    rq_activate_all_grippers(True)
    # end: URCap Program Node
  end
  $ 59 "zero_ftsensor()"
  zero_ftsensor()
  $ 60 "EXTT"
  $ 61 "Set GRP_3F_Enable=Off"
  set_standard_digital_out(4, False)
  $ 62 "Set DO[6]=Off"
  set_standard_digital_out(6, False)
  $ 63 "Set GRP_3F_Decap=Off"
  set_standard_digital_out(3, False)
  $ 64 "Set GRP_3F_Cap=Off"
  set_standard_digital_out(2, False)
  $ 65 "Set GRP_3F_Open=Off"
  set_standard_digital_out(5, False)
  $ 66 "PSE_T≔get_tool_free_pose(dir=[0,0,0.150], move_in_base_frame=True)"
  global PSE_T=get_tool_free_pose(dir=[0,0,0.150], move_in_base_frame=True)
  $ 67 "If is_reachable(Base_const, [PSE_T])"
  if (is_reachable(p[0.0,0.0,0.0,0.0,0.0,0.0], [PSE_T])):
    $ 68 "MoveL"
    $ 69 "PSE_T" "breakAfter"
    movel(PSE_T, a=1.2, v=0.15)
  end
  $ 70 "powder dispensing variable init"
  $ 71 "Start_thread≔ False "
  global Start_thread=  False
  $ 72 "vib_mot_thread≔ False "
  global vib_mot_thread=  False
  $ 73 "kp≔0.00005"
  global kp=0.00005
  $ 74 "ki≔0.0005"
  global ki=0.0005
  $ 75 "kd≔0.002"
  global kd=0.002
  $ 76 "dt≔0.02"
  global dt=0.02
  $ 77 "Integral_error≔0"
  global Integral_error=0
  $ 78 "current_error≔0"
  global current_error=0
  $ 79 "previous_error≔0"
  global previous_error=0
  $ 80 "tilt_increment≔0"
  global tilt_increment=0
  $ 81 "tilt_angle≔0"
  global tilt_angle=0
  $ 82 "diff≔0"
  global diff=0
  $ 83 "current_pose≔get_actual_tcp_pose()"
  global current_pose= get_actual_tcp_pose ()
  $ 84 "Relative_trans≔p[0, 0, -0.035, 0, 0, 0]"
  global Relative_trans=p[0, 0, -0.035, 0, 0, 0]
  $ 85 "ContA_plc_offst≔p[-0.00205, 0.02547, 0.03730, -0.03, -2.183, 6.165]"
  global ContA_plc_offst=p[-0.00205, 0.02547, 0.03730, -0.03, -2.183, 6.165]
  $ 86 "PowA_50_offset≔p[0.21808, -0.19943, 0.06584, 0, 0, 0]"
  global PowA_50_offset=p[0.21808, -0.19943, 0.06584, 0, 0, 0]
  $ 87 "scooping_init()"
  scooping_init()
  $ 88 "tilt_init_reference()"
  tilt_init_reference()
  $ 89 "switch_spatula≔ True "
  global switch_spatula=  True
  $ 679 "Thread_1"
  thread Thread_1():
    while (True):
      $ 680 "If Start_thread≟ True "
      if (Start_thread ==   True  ):
        $ 681 "Weight_value≔get_weight()"
        global Weight_value=get_weight()
        $ 682 "Wait: 0.1"
        sleep(0.1)
        $ 683 "sync()"
        sync()
      end
    end
  end
  threadId_Thread_1 = run Thread_1()
  $ 695 "Thread_2"
  thread Thread_2():
    while (True):
      $ 696 "Loop vib_mot_thread≟ True "
      thread Thread_while_696():
        while (True):
          $ 697 "diff≔Target_weight-Weight_value"
          global diff=Target_weight-Weight_value
          $ 698 "If diff>0.15"
          global thread_flag_698=0
          thread Thread_if_698():
            $ 700 "Set AO[0]=4.0"
            set_standard_analog_out(0, 0.4)
            thread_flag_698 = 1
          end
          if (diff>0.15):
            global thread_handler_698=run Thread_if_698()
            while (thread_flag_698 == 0):
              if not(diff>0.15):
                kill thread_handler_698
                thread_flag_698 = 2
              else:
                sync()
              end
            end
          else:
            thread_flag_698 = 2
          end
          if (thread_flag_698 == 2):
            $ 701 "ElseIf diff≥0.05 and diff≤0.15"
            global thread_flag_701=0
            thread Thread_if_701():
              $ 702 "vibration_2()"
              vibration_2()
              thread_flag_701 = 1
            end
            if (diff >= 0.05 and diff <= 0.15):
              global thread_handler_701=run Thread_if_701()
              while (thread_flag_701 == 0):
                if not(diff >= 0.05 and diff <= 0.15):
                  kill thread_handler_701
                  thread_flag_701 = 2
                else:
                  sync()
                end
              end
            else:
              thread_flag_701 = 2
            end
            if (thread_flag_701 == 2):
              $ 703 "ElseIf diff≥0.01 and diff<0.05"
              if (diff >= 0.01 and diff<0.05):
                $ 704 "vibration_3()"
                vibration_3()
              else:
                $ 705 "ElseIf diff>0 and diff<0.01"
                if (diff>0 and diff<0.01):
                  $ 706 "vibration_4()"
                  vibration_4()
                else:
                  $ 707 "Else" "noBreak"
                  $ 708 "Set AO[0]=0.0"
                  set_standard_analog_out(0, 0.0)
                end
              end
            end
          end
        end
      end
      if (vib_mot_thread ==   True  ):
        global thread_handler_696=run Thread_while_696()
        while (vib_mot_thread ==   True  ):
          sync()
        end
        kill thread_handler_696
      end
      $ 712 "sync()"
      sync()
    end
  end
  threadId_Thread_2 = run Thread_2()
  while (True):
    $ 90 "Robot Program"
    $ 91 "MAIN"
    $ 92 "command_manager(external_control='uGO', cond_suspend=(ITM_Manipulated and AMR_AtTarget and AMR_Charging and AMR_Battery<40), cond_unsuspend=(AMR_Battery≟60))"
    command_manager(external_control="uGO", cond_suspend=(ITM_Manipulated  and  AMR_AtTarget  and  AMR_Charging  and  AMR_Battery<40), cond_unsuspend=(AMR_Battery == 60))
    $ 93 "log_state(STATE_Info)"
    log_state(STATE_Info)
    $ 94 "Switch STATE"
    switch_1 = STATE
    $ 95 "Case 1"
    if (1 == switch_1):
      $ 96 "Stopping"
      $ 97 "STATE_Info≔'Stopping'"
      global STATE_Info="Stopping"
      $ 98 "end_freedrive_mode()"
      end_freedrive_mode()
      $ 99 "Set"
      set_tcp(p[0.0,0.0,0.161,3.1415,0.0,0.0])
      $ 100 "PSE_T≔get_tool_free_pose(dir=[0,0,0.150], move_in_base_frame=True)"
      global PSE_T=get_tool_free_pose(dir=[0,0,0.150], move_in_base_frame=True)
      $ 101 "If is_reachable(Base_const, [PSE_T])"
      if (is_reachable(p[0.0,0.0,0.0,0.0,0.0,0.0], [PSE_T])):
        $ 102 "MoveL"
        $ 103 "PSE_T" "breakAfter"
        movel(PSE_T, a=1.2, v=0.15)
      end
      $ 104 "do_transition(keep_rxry=OBJ_Picked, r=0)"
      do_transition(keep_rxry=OBJ_Picked, r=0)
      $ 113 "Call Sub_AMR_MiR_V3"
      Sub_AMR_MiR_V3()
      $ 114 "If stopping() and AMR_Done"
      if (stopping()  and  AMR_Done):
        $ 115 "STATE≔2"
        global STATE=2
        $ 116 "ugo_update_outputs()"
        ugo_update_outputs()
      end
    elif (2 == switch_1):
      $ 117 "Case 2"
      $ 118 "Stopped"
      $ 119 "STATE_Info≔'Stopped'"
      global STATE_Info="Stopped"
      $ 120 "Call Sub_AMR_MiR_V3"
      Sub_AMR_MiR_V3()
      $ 121 "If CMD_Reset"
      if (CMD_Reset):
        $ 122 "STATE≔3"
        global STATE=3
        $ 123 "ugo_update_outputs()"
        ugo_update_outputs()
      end
    elif (3 == switch_1):
      $ 124 "Case 3"
      $ 125 " Resetting"
      $ 126 "STATE_Info≔'Resetting'"
      global STATE_Info="Resetting"
      $ 127 "uML"
      $ 128 "reset_error()"
      reset_error()
      $ 129 "reset_warning()"
      reset_warning()
      $ 130 "PROCESS_Step≔0"
      global PROCESS_Step=0
      $ 131 "PROCESS_Info≔''"
      global PROCESS_Info=""
      $ 132 "ARM_Referenced≔ False "
      global ARM_Referenced=  False
      $ 133 "WRK_Done≔ False "
      global WRK_Done=  False
      $ 134 "ITM_Prepared≔ False "
      global ITM_Prepared=  False
      $ 135 "ITM_Manipulated≔ False "
      global ITM_Manipulated=  False
      $ 136 "STP≔0"
      global STP=0
      $ 137 "Action≔0"
      global Action=0
      $ 138 "Action_Info≔''"
      global Action_Info=""
      $ 139 "ITM_ID≔0"
      global ITM_ID=0
      $ 140 "JIG≔0"
      global JIG=0
      $ 141 "JIG_Slot≔0"
      global JIG_Slot=0
      $ 142 "Task_info≔''"
      global Task_info=""
      $ 143 "Set"
      set_tcp(p[0.0,0.0,0.161,3.1415,0.0,0.0])
      $ 144 "App"
      $ 145 "'ADD APPLICATION SPECIFIC COMMANDS'"
      # 'ADD APPLICATION SPECIFIC COMMANDS'
      $ 146 "OBJ_Type≔0"
      global OBJ_Type=0
      $ 147 "OBJ_Nbr≔0"
      global OBJ_Nbr=0
      $ 148 "If CNT_Rack_Output≥50"
      if (CNT_Rack_Output >= 50):
        $ 149 "CNT_Rack_Output≔0"
        global CNT_Rack_Output=0
      end
      $ 150 "TASK≔struct(ID=0, NAVI=struct(target=0, footprint=0, protectiveOff=0, dock=0), WORK=struct(ITM_ID_Src=0, JIG_ID_Src=0, OBJ_Nbr_Src=0, ACT_Src=0, ITM_ID_Tgt=0, JIG_ID_Tgt=0, OBJ_Nbr_Tgt=0, ACT_Tgt=0, OBJ_Type=0))"
      global TASK=struct(ID=0, NAVI=struct(target=0, footprint=0, protectiveOff=0, dock=0), WORK=struct(ITM_ID_Src=0, JIG_ID_Src=0, OBJ_Nbr_Src=0, ACT_Src=0, ITM_ID_Tgt=0, JIG_ID_Tgt=0, OBJ_Nbr_Tgt=0, ACT_Tgt=0, OBJ_Type=0))
      $ 151 "Call Sub_AMR_MiR_V3"
      Sub_AMR_MiR_V3()
      $ 152 "If resetting() and AMR_Done"
      if (resetting()  and  AMR_Done):
        $ 153 "STATE≔4"
        global STATE=4
        $ 154 "ugo_update_outputs()"
        ugo_update_outputs()
      end
    elif (4 == switch_1):
      $ 155 "Case 4"
      $ 156 "Idle"
      $ 157 "STATE_Info≔'Idle'"
      global STATE_Info="Idle"
      $ 158 "If CMD_Start"
      if (CMD_Start):
        $ 159 "STATE≔5"
        global STATE=5
        $ 160 "ugo_update_outputs()"
        ugo_update_outputs()
      end
    elif (5 == switch_1):
      $ 161 "Case 5"
      $ 162 "Starting"
      $ 163 "STATE_Info≔'Starting'"
      global STATE_Info="Starting"
      $ 164 "'ADD COMMANDS WHAT TO START WITH'"
      # 'ADD COMMANDS WHAT TO START WITH'
      $ 165 "Call Sub_AMR_MiR_V3"
      Sub_AMR_MiR_V3()
      $ 166 "get ugo data"
      $ 167 "Assign Tasks"
      $ 168 "TASK.ID = ugo_get_task()"
      TASK.ID = ugo_get_task()
      $ 169 "If TASK.ID≟1"
      if (TASK.ID == 1):
        $ 170 "Task_info≔'Charge'"
        global Task_info="Charge"
        $ 171 "Parameters"
        $ 172 "AMR_PosTarget≔1"
        global AMR_PosTarget=1
      else:
        $ 173 "ElseIf TASK.ID≟9"
        if (TASK.ID == 9):
          $ 174 "'Pick Sarstedt Rack from Variable source'"
          # 'Pick Sarstedt Rack from Variable source'
          $ 175 "Task_info≔'Navigate to Target'"
          global Task_info="Navigate to Target"
          $ 176 "Parameters"
          $ 177 "AMR_PosTarget≔UGO.read_input('00','ITM_ID')"
          global AMR_PosTarget=UGO.read_input("00","ITM_ID")
        else:
          $ 178 "ElseIf TASK.ID≟49"
          if (TASK.ID == 49):
            $ 179 "Task_info≔'Pick Containers'"
            global Task_info="Pick Containers"
            $ 180 "Parameters"
            $ 181 "ITM_ID≔1"
            global ITM_ID=1
            $ 182 "OBJ_Type≔6"
            global OBJ_Type=6
            $ 183 "JIG≔15"
            global JIG=15
            $ 184 "AMR_PosTarget≔3"
            global AMR_PosTarget=3
          else:
            $ 185 "ElseIf TASK.ID≟50"
            if (TASK.ID == 50):
              $ 186 "Task_info≔'Decap Containers'"
              global Task_info="Decap Containers"
              $ 187 "Parameters"
              $ 188 "ITM_ID≔1"
              global ITM_ID=1
              $ 189 "OBJ_Type≔6"
              global OBJ_Type=6
              $ 190 "JIG≔16"
              global JIG=16
              $ 191 "AMR_PosTarget≔5"
              global AMR_PosTarget=5
            else:
              $ 192 "ElseIf TASK.ID≟51"
              if (TASK.ID == 51):
                $ 193 "Task_info≔'Detect Spatula and transfer powder'"
                global Task_info="Detect Spatula and transfer powder"
                $ 194 "Parameters"
                $ 195 "ITM_ID≔1"
                global ITM_ID=1
                $ 196 "Target_weight≔(UGO.read_input('00','Target_weight'))/1000"
                global Target_weight=(UGO.read_input("00","Target_weight"))/1000
                $ 197 "OBJ_Type≔8"
                global OBJ_Type=8
                $ 198 "JIG≔16"
                global JIG=16
                $ 199 "AMR_PosTarget≔5"
                global AMR_PosTarget=5
              else:
                $ 200 "ElseIf TASK.ID≟52"
                if (TASK.ID == 52):
                  $ 201 "Task_info≔'Pick PowderA'"
                  global Task_info="Pick PowderA"
                  $ 202 "Parameters"
                  $ 203 "ITM_ID≔1"
                  global ITM_ID=1
                  $ 204 "OBJ_Type≔6"
                  global OBJ_Type=6
                  $ 205 "JIG≔15"
                  global JIG=15
                  $ 206 "AMR_PosTarget≔3"
                  global AMR_PosTarget=3
                else:
                  $ 207 "ElseIf TASK.ID≟53"
                  if (TASK.ID == 53):
                    $ 208 "Task_info≔'Decap PowderA'"
                    global Task_info="Decap PowderA"
                    $ 209 "Parameters"
                    $ 210 "ITM_ID≔1"
                    global ITM_ID=1
                    $ 211 "OBJ_Type≔6"
                    global OBJ_Type=6
                    $ 212 "JIG≔1"
                    global JIG=1
                    $ 213 "AMR_PosTarget≔5"
                    global AMR_PosTarget=5
                  else:
                    $ 214 "ElseIf TASK.ID≟54"
                    if (TASK.ID == 54):
                      $ 215 "Task_info≔'Dispense PowderA'"
                      global Task_info="Dispense PowderA"
                      $ 216 "Parameters"
                      $ 217 "ITM_ID≔1"
                      global ITM_ID=1
                      $ 218 "Target_weight≔(UGO.read_input('00','Target_weight'))/1000"
                      global Target_weight=(UGO.read_input("00","Target_weight"))/1000
                      $ 219 "W_now≔(UGO.read_input('00','Container_weight'))/1000"
                      global W_now=(UGO.read_input("00","Container_weight"))/1000
                      $ 220 "Powder_name≔(UGO.read_input('00','Powder_name'))"
                      global Powder_name=(UGO.read_input("00","Powder_name"))
                      $ 221 "OBJ_Type≔6"
                      global OBJ_Type=6
                      $ 222 "JIG≔17"
                      global JIG=17
                      $ 223 "AMR_PosTarget≔5"
                      global AMR_PosTarget=5
                    else:
                      $ 224 "ElseIf TASK.ID≟55"
                      if (TASK.ID == 55):
                        $ 225 "Task_info≔'Place PowderA'"
                        global Task_info="Place PowderA"
                        $ 226 "Parameters"
                        $ 227 "ITM_ID≔1"
                        global ITM_ID=1
                        $ 228 "OBJ_Type≔6"
                        global OBJ_Type=6
                        $ 229 "JIG≔21"
                        global JIG=21
                        $ 230 "AMR_PosTarget≔5"
                        global AMR_PosTarget=5
                      else:
                        $ 231 "Else" "noBreak"
                        $ 232 "set_error(ERROR_WRONG_ORDER)"
                        set_error(ERROR_WRONG_ORDER)
                      end
                    end
                  end
                end
              end
            end
          end
        end
      end
      $ 233 "test ugo"
      $ 234 "Wait: 0.2"
      sleep(0.2)
      $ 235 "ugo_update_outputs()"
      ugo_update_outputs()
      $ 236 "If starting() and AMR_Done"
      if (starting()  and  AMR_Done):
        $ 237 "log_message(Task_info, 'New Task: ')"
        log_message(Task_info, "New Task: ")
        $ 238 "log_message(to_str(TASK.ID), 'Task_ID: ')"
        log_message(to_str(TASK.ID), "Task_ID: ")
        $ 239 "do_transition(keep_rxry=OBJ_Picked)"
        do_transition(keep_rxry=OBJ_Picked)
        $ 240 "STATE≔6"
        global STATE=6
        $ 241 "ugo_update_outputs()"
        ugo_update_outputs()
      end
    elif (6 == switch_1):
      $ 242 "Case 6"
      $ 243 "Execute"
      $ 244 "STATE_Info≔'Execute'"
      global STATE_Info="Execute"
      $ 245 "If  not CMD_Hold and not CMD_Suspend"
      global thread_flag_245=0
      thread Thread_if_245():
        $ 246 "Switch PROCESS_Step"
        switch_2 = PROCESS_Step
        $ 247 "Case 0"
        if (0 == switch_2):
          $ 248 "PROCESS_Info≔'process control'"
          global PROCESS_Info="process control"
          $ 249 "log_process(PROCESS_Info)"
          log_process(PROCESS_Info)
          $ 250 "process control"
          $ 251 "If  not AMR_AtTarget"
          if (  not  AMR_AtTarget):
            $ 252 "PROCESS_Step≔1"
            global PROCESS_Step=1
          else:
            $ 253 "ElseIf (( not ITM_Prepared and  not WRK_Done) or (ITM_Prepared and WRK_Done))"
            if (((  not  ITM_Prepared  and    not  WRK_Done)  or  (ITM_Prepared  and  WRK_Done))):
              $ 254 "PROCESS_Step≔2"
              global PROCESS_Step=2
            else:
              $ 255 "ElseIf  not WRK_Done"
              if (  not  WRK_Done):
                $ 256 "PROCESS_Step≔3"
                global PROCESS_Step=3
              else:
                $ 257 "Else" "noBreak"
                $ 258 "task finished"
                $ 259 "PROCESS_Info≔''"
                global PROCESS_Info=""
                $ 260 "STATE≔7"
                global STATE=7
                $ 261 "ugo_update_outputs()"
                ugo_update_outputs()
              end
            end
          end
        elif (1 == switch_2):
          $ 262 "Case 1"
          $ 263 "navigate"
          $ 264 "'MOVING THE uML'"
          # 'MOVING THE uML'
          $ 265 "PROCESS_Info≔'move to target'"
          global PROCESS_Info="move to target"
          $ 266 "log_process(PROCESS_Info)"
          log_process(PROCESS_Info)
          $ 267 "If TASK.ID≟1"
          if (TASK.ID == 1):
            $ 268 "Action≔51"
            global Action=51
          else:
            $ 269 "Else" "noBreak"
            $ 270 "Action≔52"
            global Action=52
          end
          $ 271 "Call Sub_AMR_MiR_V3"
          Sub_AMR_MiR_V3()
          $ 272 "If AMR_Done"
          if (AMR_Done):
            $ 273 "PROCESS_Step≔0"
            global PROCESS_Step=0
          end
        elif (2 == switch_2):
          $ 274 "Case 2"
          $ 275 "prepare"
          $ 276 "'THINGS THAT HAVE TO BE DONE ONCE IN A SEQUENCE,WORKFLOW'"
          # 'THINGS THAT HAVE TO BE DONE ONCE IN A SEQUENCE,WORKFLOW'
          $ 277 "PROCESS_Info≔'prepare for work'"
          global PROCESS_Info="prepare for work"
          $ 278 "log_process(PROCESS_Info)"
          log_process(PROCESS_Info)
          $ 279 "If TASK.WORK.ITM_ID_Src>1"
          if (TASK.WORK.ITM_ID_Src>1):
            $ 280 "ITM_ID≔TASK.WORK.ITM_ID_Src"
            global ITM_ID=TASK.WORK.ITM_ID_Src
          else:
            $ 281 "ElseIf TASK.WORK.ITM_ID_Tgt>1"
            if (TASK.WORK.ITM_ID_Tgt>1):
              $ 282 "ITM_ID≔TASK.WORK.ITM_ID_Tgt"
              global ITM_ID=TASK.WORK.ITM_ID_Tgt
            end
          end
          $ 283 "If  not ARM_Referenced and (ITM_ID≠0)"
          if (  not  ARM_Referenced  and  (ITM_ID != 0)):
            $ 284 "STP≔1"
            global STP=1
          else:
            $ 285 "ElseIf ARM_Referenced or (ITM_ID≟0)"
            if (ARM_Referenced  or  (ITM_ID == 0)):
              $ 286 "STP≔2"
              global STP=2
            end
          end
          $ 287 "Switch STP"
          switch_3 = STP
          $ 288 "Case 1"
          if (1 == switch_3):
            $ 289 "reference"
            $ 290 "STP_Info≔'reference at target position'"
            global STP_Info="reference at target position"
            $ 291 "log_step(STP_Info)"
            log_step(STP_Info)
            $ 292 "If ITM_ID≟1"
            if (ITM_ID == 1):
              $ 293 "CAM_Done≔ True "
              global CAM_Done=  True
            else:
              $ 294 "Else" "noBreak"
              $ 295 "Action≔131"
              global Action=131
              $ 296 "Call Sub_Vision_V18"
              Sub_Vision_V18()
            end
            $ 298 "If CAM_Done and  not ERROR.FLAG"
            if (CAM_Done  and    not  ERROR.FLAG):
              $ 299 "log_step('ARM referenced')"
              log_step("ARM referenced")
              $ 300 "ARM_Referenced≔ True "
              global ARM_Referenced=  True
            end
          elif (2 == switch_3):
            $ 301 "Case 2"
            $ 302 "manipulate"
            $ 303 "STP_Info≔'manipulate item'"
            global STP_Info="manipulate item"
            $ 304 "log_step(STP_Info)"
            log_step(STP_Info)
            $ 305 "'In case pressing button is needed'"
            # 'In case pressing button is needed'
            $ 306 "If found_in_list(ITM_ID, ITM_ID_List)"
            if (found_in_list(ITM_ID, ITM_ID_List)):
              $ 307 "Switch ITM_ID"
              switch_4 = ITM_ID
              $ 308 "Case 0"
              if (0 == switch_4):
                $ 309 "ITM_Manipulated≔ not ITM_Manipulated"
                global ITM_Manipulated=  not  ITM_Manipulated
              elif (1 == switch_4):
                $ 310 "Case 1"
                $ 311 "ITM_Manipulated≔ not ITM_Manipulated"
                global ITM_Manipulated=  not  ITM_Manipulated
              elif (2 == switch_4):
                $ 312 "Case 2"
              else:
                $ 322 "Default Case"
                $ 323 "ITM_Manipulated≔ not ITM_Manipulated"
                global ITM_Manipulated=  not  ITM_Manipulated
              end
            end
          end
          $ 324 "ITM_Prepared≔(ITM_Manipulated or  not found_in_list(ITM_ID, ITM_ID_List)) and (ARM_Referenced or ITM_ID≟0) and  not WRK_Done"
          global ITM_Prepared=(ITM_Manipulated  or    not  found_in_list(ITM_ID, ITM_ID_List))  and  (ARM_Referenced  or  ITM_ID == 0)  and    not  WRK_Done
          $ 325 "STP≔0"
          global STP=0
          $ 326 "STP_Info≔''"
          global STP_Info=""
          $ 327 "PROCESS_Step≔0"
          global PROCESS_Step=0
        elif (3 == switch_2):
          $ 328 "Case 3"
          $ 329 "work"
          $ 330 "'ADD EVERY MACHINE, OBJECT, STATION TO WORK ON'"
          # 'ADD EVERY MACHINE, OBJECT, STATION TO WORK ON'
          $ 331 "Switch ITM_ID"
          switch_3 = ITM_ID
          $ 332 "Case 1"
          if (1 == switch_3):
            $ 333 "uLM"
            $ 334 "If TASK.ID≟12"
            if (TASK.ID == 12):
              $ 335 "fill racks"
              $ 336 "Action≔151"
              global Action=151
              $ 337 "Call Sub_Vision_V18"
              Sub_Vision_V18()
              $ 338 "If  not ERROR.FLAG"
              if (  not  ERROR.FLAG):
                $ 339 "Actions for the task"
                $ 340 "Action≔1"
                global Action=1
                $ 341 "JIG≔2"
                global JIG=2
                $ 342 "JIG_Slot≔CAM_Result[0]"
                global JIG_Slot=CAM_Result[0]
                $ 343 "OBJ_Nbr≔CAM_Result[0]"
                global OBJ_Nbr=CAM_Result[0]
                $ 344 "OBJ_Type≔2"
                global OBJ_Type=2
                $ 345 "Call Sub_Action_V4"
                Sub_Action_V4()
                $ 346 "If OBJ_Picked"
                if (OBJ_Picked):
                  $ 347 "CAM_Result.remove(0)"
                  CAM_Result.remove(0)
                  $ 348 "PRC_TubCounter≔PRC_TubCounter+1"
                  global PRC_TubCounter=PRC_TubCounter+1
                  $ 349 "If PRC_TubCounter%4≟0"
                  if (PRC_TubCounter%4 == 0):
                    $ 350 "JIG_Slot≔4"
                    global JIG_Slot=4
                  else:
                    $ 351 "Else" "noBreak"
                    $ 352 "JIG_Slot≔PRC_TubCounter%4"
                    global JIG_Slot=PRC_TubCounter%4
                  end
                  $ 353 "OBJ_Nbr≔ceil(PRC_TubCounter/4)"
                  global OBJ_Nbr=ceil(PRC_TubCounter/4)
                  $ 354 "Action≔2"
                  global Action=2
                  $ 355 "JIG≔4"
                  global JIG=4
                  $ 356 "Call Sub_Action_V4"
                  Sub_Action_V4()
                  $ 357 "Action≔151"
                  global Action=151
                  $ 358 "Call Sub_Vision_V18"
                  Sub_Vision_V18()
                end
              end
              $ 359 "If (CAM_Captures≥CAM_PRM_Retries) or (PRC_TubCounter≥32)"
              if ((CAM_Captures >= CAM_PRM_Retries)  or  (PRC_TubCounter >= 32)):
                $ 360 "PROCESS_Step≔0"
                global PROCESS_Step=0
                $ 361 "WRK_Done≔ True "
                global WRK_Done=  True
              end
            else:
              $ 362 "ElseIf TASK.ID≟49"
              if (TASK.ID == 49):
                $ 363 "Pick Powder container"
                $ 364 "Action≔131"
                global Action=131
                $ 365 "Call Sub_Vision_V18"
                Sub_Vision_V18()
                $ 366 "Action≔35"
                global Action=35
                $ 367 "Call Sub_Action_V4"
                Sub_Action_V4()
                $ 368 "PROCESS_Step≔0"
                global PROCESS_Step=0
                $ 369 "WRK_Done≔ True "
                global WRK_Done=  True
              else:
                $ 370 "ElseIf TASK.ID≟50"
                if (TASK.ID == 50):
                  $ 371 "Decap containers"
                  $ 372 "Action≔36"
                  global Action=36
                  $ 373 "Call Sub_Action_V4"
                  Sub_Action_V4()
                  $ 374 "PROCESS_Step≔0"
                  global PROCESS_Step=0
                  $ 375 "WRK_Done≔ True "
                  global WRK_Done=  True
                else:
                  $ 376 "ElseIf TASK.ID≟51"
                  if (TASK.ID == 51):
                    $ 377 "Detect Spatula and transfer powder"
                    $ 378 "Action≔131"
                    global Action=131
                    $ 379 "Call Sub_Vision_V18"
                    Sub_Vision_V18()
                    $ 380 "Action≔37"
                    global Action=37
                    $ 381 "Call Sub_Action_V4"
                    Sub_Action_V4()
                    $ 382 "PROCESS_Step≔0"
                    global PROCESS_Step=0
                    $ 383 "WRK_Done≔ True "
                    global WRK_Done=  True
                  else:
                    $ 384 "ElseIf TASK.ID≟52"
                    if (TASK.ID == 52):
                      $ 385 "Pick PowderA container"
                      $ 386 "Action≔131"
                      global Action=131
                      $ 387 "Call Sub_Vision_V18"
                      Sub_Vision_V18()
                      $ 388 "Action≔38"
                      global Action=38
                      $ 389 "Call Sub_Action_V4"
                      Sub_Action_V4()
                      $ 390 "PROCESS_Step≔0"
                      global PROCESS_Step=0
                      $ 391 "WRK_Done≔ True "
                      global WRK_Done=  True
                    else:
                      $ 392 "ElseIf TASK.ID≟53"
                      if (TASK.ID == 53):
                        $ 393 "Decap containerA"
                        $ 394 "Action≔39"
                        global Action=39
                        $ 395 "Call Sub_Action_V4"
                        Sub_Action_V4()
                        $ 396 "PROCESS_Step≔0"
                        global PROCESS_Step=0
                        $ 397 "WRK_Done≔ True "
                        global WRK_Done=  True
                      else:
                        $ 398 "ElseIf TASK.ID≟55"
                        if (TASK.ID == 55):
                          $ 399 "Place PowderA"
                          $ 400 "Action≔131"
                          global Action=131
                          $ 401 "Call Sub_Vision_V18"
                          Sub_Vision_V18()
                          $ 402 "Action≔40"
                          global Action=40
                          $ 403 "Call Sub_Action_V4"
                          Sub_Action_V4()
                          $ 404 "PROCESS_Step≔0"
                          global PROCESS_Step=0
                          $ 405 "WRK_Done≔ True "
                          global WRK_Done=  True
                        else:
                          $ 406 "ElseIf TASK.ID≟54"
                          if (TASK.ID == 54):
                            $ 407 "Dispense PowderA"
                            $ 408 "Action≔131"
                            global Action=131
                            $ 409 "Call Sub_Vision_V18"
                            Sub_Vision_V18()
                            $ 410 "Action≔41"
                            global Action=41
                            $ 411 "Call Sub_Action_V4"
                            Sub_Action_V4()
                            $ 412 "PROCESS_Step≔0"
                            global PROCESS_Step=0
                            $ 413 "WRK_Done≔ True "
                            global WRK_Done=  True
                          end
                        end
                      end
                    end
                  end
                end
              end
            end
          elif (2 == switch_3):
            $ 414 "Case 2"
          elif (5 == switch_3):
            $ 456 "Case 5"
          elif (20 == switch_3):
            $ 464 "Case 20"
          elif (43 == switch_3):
            $ 526 "Case 43"
          else:
            $ 534 "Default Case"
            $ 535 "WRK_Done≔ True "
            global WRK_Done=  True
            $ 536 "PROCESS_Step≔0"
            global PROCESS_Step=0
          end
        end
        thread_flag_245 = 1
      end
      if (  not  CMD_Hold and not CMD_Suspend):
        global thread_handler_245=run Thread_if_245()
        while (thread_flag_245 == 0):
          if not(  not  CMD_Hold and not CMD_Suspend):
            kill thread_handler_245
            thread_flag_245 = 2
          else:
            sync()
          end
        end
      else:
        thread_flag_245 = 2
      end
      $ 537 "If CMD_Hold"
      if (CMD_Hold):
        $ 538 "STATE≔9"
        global STATE=9
        $ 539 "ugo_update_outputs()"
        ugo_update_outputs()
      else:
        $ 540 "ElseIf CMD_Suspend"
        if (CMD_Suspend):
          $ 541 "STATE≔12"
          global STATE=12
          $ 542 "ugo_update_outputs()"
          ugo_update_outputs()
        end
      end
    elif (7 == switch_1):
      $ 543 "Case 7"
      $ 544 "Completing"
      $ 545 "STATE_Info≔'Completing'"
      global STATE_Info="Completing"
      $ 546 "'ADD COMMANDS FOR COMPLETING THE PROCESS'"
      # 'ADD COMMANDS FOR COMPLETING THE PROCESS'
      $ 547 "do_transition(keep_rxry=OBJ_Picked)"
      do_transition(keep_rxry=OBJ_Picked)
      $ 548 "Call Sub_AMR_MiR_V3"
      Sub_AMR_MiR_V3()
      $ 549 "If completing() and AMR_Done"
      if (completing()  and  AMR_Done):
        $ 550 "STATE≔8"
        global STATE=8
        $ 551 "ugo_update_outputs()"
        ugo_update_outputs()
      end
    elif (8 == switch_1):
      $ 552 "Case 8"
      $ 553 "Complete"
      $ 554 "STATE_Info≔'Complete'"
      global STATE_Info="Complete"
      $ 555 "If CMD_Reset"
      if (CMD_Reset):
        $ 556 "STATE≔3"
        global STATE=3
        $ 557 "ugo_update_outputs()"
        ugo_update_outputs()
      end
    elif (9 == switch_1):
      $ 558 "Case 9"
      $ 559 "Holding"
      $ 560 "STATE_Info≔'Holding'"
      global STATE_Info="Holding"
      $ 561 "stopl(0.5)"
      stopl(0.5)
      $ 562 "Call Sub_AMR_MiR_V3"
      Sub_AMR_MiR_V3()
      $ 563 "If holding() and AMR_Done"
      if (holding()  and  AMR_Done):
        $ 564 "STATE≔10"
        global STATE=10
        $ 565 "ugo_update_outputs()"
        ugo_update_outputs()
      end
    elif (10 == switch_1):
      $ 566 "Case 10"
      $ 567 "Held"
      $ 568 "STATE_Info≔'Held'"
      global STATE_Info="Held"
      $ 569 "If CMD_Unhold"
      if (CMD_Unhold):
        $ 570 "end_freedrive_mode()"
        end_freedrive_mode()
        $ 571 "STATE≔11"
        global STATE=11
        $ 572 "ugo_update_outputs()"
        ugo_update_outputs()
      else:
        $ 573 "ElseIf FNC_Freedrive"
        if (FNC_Freedrive):
          $ 574 "freedrive_mode()"
          freedrive_mode()
        else:
          $ 575 "Else" "noBreak"
          $ 576 "end_freedrive_mode()"
          end_freedrive_mode()
        end
      end
    elif (11 == switch_1):
      $ 577 "Case 11"
      $ 578 "Unholding"
      $ 579 "STATE_Info≔'Unholding'"
      global STATE_Info="Unholding"
      $ 580 "Clearing"
      $ 581 "Switch ERROR.ID"
      switch_2 = ERROR.ID
      $ 582 "Case 1002"
      if (1002 == switch_2):
        $ 583 "AMR_AtTarget≔ False "
        global AMR_AtTarget=  False
        $ 584 "ARM_Referenced≔ False "
        global ARM_Referenced=  False
        $ 585 "ITM_Prepared≔ False "
        global ITM_Prepared=  False
        $ 586 "PROCESS_Step≔1"
        global PROCESS_Step=1
      elif (2007 == switch_2):
        $ 587 "Case 2007"
        $ 588 "PROCESS_Step≔1"
        global PROCESS_Step=1
      end
      $ 589 "reset_error()"
      reset_error()
      $ 590 "reset_warning()"
      reset_warning()
      $ 591 "OBJ_Picked≔gripper_has_object()"
      global OBJ_Picked=gripper_has_object()
      $ 592 "Call Sub_AMR_MiR_V3"
      Sub_AMR_MiR_V3()
      $ 593 "If unholding() and AMR_Done"
      if (unholding()  and  AMR_Done):
        $ 594 "STATE≔6"
        global STATE=6
        $ 595 "ugo_update_outputs()"
        ugo_update_outputs()
      end
    elif (12 == switch_1):
      $ 596 "Case 12"
      $ 597 "Suspending"
      $ 598 "STATE_Info≔'Suspending'"
      global STATE_Info="Suspending"
      $ 599 "PROCESS_Info≔str_cat(PROCESS_Info, ' suspended')"
      global PROCESS_Info=str_cat(PROCESS_Info, " suspended")
      $ 600 "If suspending()"
      if (suspending()):
        $ 601 "STATE≔13"
        global STATE=13
        $ 602 "ugo_update_outputs()"
        ugo_update_outputs()
      end
    elif (13 == switch_1):
      $ 603 "Case 13"
      $ 604 "Suspended"
      $ 605 "STATE_Info≔'Suspended'"
      global STATE_Info="Suspended"
      $ 606 "Call Sub_AMR_MiR_V3"
      Sub_AMR_MiR_V3()
      $ 607 "If CMD_Unsuspend"
      if (CMD_Unsuspend):
        $ 608 "STATE≔14"
        global STATE=14
        $ 609 "ugo_update_outputs()"
        ugo_update_outputs()
      end
    elif (14 == switch_1):
      $ 610 "Case 14"
      $ 611 "Unsuspending"
      $ 612 "STATE_Info≔'Unsuspending'"
      global STATE_Info="Unsuspending"
      $ 613 "PROCESS_Step≔0"
      global PROCESS_Step=0
      $ 614 "If unsuspending()"
      if (unsuspending()):
        $ 615 "STATE≔6"
        global STATE=6
        $ 616 "ugo_update_outputs()"
        ugo_update_outputs()
      end
    elif (15 == switch_1):
      $ 617 "Case 15"
      $ 618 "Aborting"
      $ 619 "STATE_Info≔'Aborting'"
      global STATE_Info="Aborting"
      $ 620 "If aborting()"
      if (aborting()):
        $ 621 "STATE≔16"
        global STATE=16
        $ 622 "ugo_update_outputs()"
        ugo_update_outputs()
      end
    elif (16 == switch_1):
      $ 623 "Case 16"
      $ 624 "Aborted"
      $ 625 "STATE_Info≔'Aborted'"
      global STATE_Info="Aborted"
      $ 626 "If CMD_Clear"
      if (CMD_Clear):
        $ 627 "STATE≔17"
        global STATE=17
        $ 628 "ugo_update_outputs()"
        ugo_update_outputs()
      end
    elif (17 == switch_1):
      $ 629 "Case 17"
      $ 630 "Clearing"
      $ 631 "STATE_Info≔'Clearing'"
      global STATE_Info="Clearing"
      $ 632 "Clearing"
      $ 633 "reset_warning()"
      reset_warning()
      $ 634 "reset_error()"
      reset_error()
      $ 635 "If clearing()"
      if (clearing()):
        $ 636 "STATE≔2"
        global STATE=2
        $ 637 "ugo_update_outputs()"
        ugo_update_outputs()
      end
    end
    $ 638 "log_state(STATE_Info)"
    log_state(STATE_Info)
    $ 639 "log_warning(WARNING.MSG)"
    log_warning(WARNING.MSG)
    $ 640 "log_error(ERROR.MSG)"
    log_error(ERROR.MSG)
    $ 641 "Times"
    $ 642 "Switch STATE"
    switch_1 = STATE
    $ 643 "Case 1"
    if (1 == switch_1):
      $ 644 "TM_St_Stopping≔get_time(STATE_Times[STATE-1])"
      global TM_St_Stopping=get_time(STATE_Times[STATE-1])
    elif (2 == switch_1):
      $ 645 "Case 2"
      $ 646 "TM_St_Stopped≔get_time(STATE_Times[STATE-1])"
      global TM_St_Stopped=get_time(STATE_Times[STATE-1])
    elif (3 == switch_1):
      $ 647 "Case 3"
      $ 648 "TM_St_Resetting≔get_time(STATE_Times[STATE-1])"
      global TM_St_Resetting=get_time(STATE_Times[STATE-1])
    elif (4 == switch_1):
      $ 649 "Case 4"
      $ 650 "TM_St_Idle≔get_time(STATE_Times[STATE-1])"
      global TM_St_Idle=get_time(STATE_Times[STATE-1])
    elif (5 == switch_1):
      $ 651 "Case 5"
      $ 652 "TM_St_Starting≔get_time(STATE_Times[STATE-1])"
      global TM_St_Starting=get_time(STATE_Times[STATE-1])
    elif (6 == switch_1):
      $ 653 "Case 6"
      $ 654 "TM_St_Execute≔get_time(STATE_Times[STATE-1])"
      global TM_St_Execute=get_time(STATE_Times[STATE-1])
    elif (7 == switch_1):
      $ 655 "Case 7"
      $ 656 "TM_St_Completin≔get_time(STATE_Times[STATE-1])"
      global TM_St_Completin=get_time(STATE_Times[STATE-1])
    elif (8 == switch_1):
      $ 657 "Case 8"
      $ 658 "TM_St_Complete≔get_time(STATE_Times[STATE-1])"
      global TM_St_Complete=get_time(STATE_Times[STATE-1])
    elif (9 == switch_1):
      $ 659 "Case 9"
      $ 660 "TM_St_Holding≔get_time(STATE_Times[STATE-1])"
      global TM_St_Holding=get_time(STATE_Times[STATE-1])
    elif (10 == switch_1):
      $ 661 "Case 10"
      $ 662 "TM_St_Held≔get_time(STATE_Times[STATE-1])"
      global TM_St_Held=get_time(STATE_Times[STATE-1])
    elif (11 == switch_1):
      $ 663 "Case 11"
      $ 664 "TM_St_Unholding≔get_time(STATE_Times[STATE-1])"
      global TM_St_Unholding=get_time(STATE_Times[STATE-1])
    elif (12 == switch_1):
      $ 665 "Case 12"
      $ 666 "TM_St_Suspendin≔get_time(STATE_Times[STATE-1])"
      global TM_St_Suspendin=get_time(STATE_Times[STATE-1])
    elif (13 == switch_1):
      $ 667 "Case 13"
      $ 668 "TM_St_Suspended≔get_time(STATE_Times[STATE-1])"
      global TM_St_Suspended=get_time(STATE_Times[STATE-1])
    elif (14 == switch_1):
      $ 669 "Case 14"
      $ 670 "TM_St_Unsuspend≔get_time(STATE_Times[STATE-1])"
      global TM_St_Unsuspend=get_time(STATE_Times[STATE-1])
    elif (15 == switch_1):
      $ 671 "Case 15"
      $ 672 "TM_St_Aborting≔get_time(STATE_Times[STATE-1])"
      global TM_St_Aborting=get_time(STATE_Times[STATE-1])
    elif (16 == switch_1):
      $ 673 "Case 16"
      $ 674 "TM_St_Aborted≔get_time(STATE_Times[STATE-1])"
      global TM_St_Aborted=get_time(STATE_Times[STATE-1])
    elif (17 == switch_1):
      $ 675 "Case 17"
      $ 676 "TM_St_Clearing≔get_time(STATE_Times[STATE-1])"
      global TM_St_Clearing=get_time(STATE_Times[STATE-1])
    end
    $ 678 "Wait: 0.1"
    sleep(0.1)
  end
end
